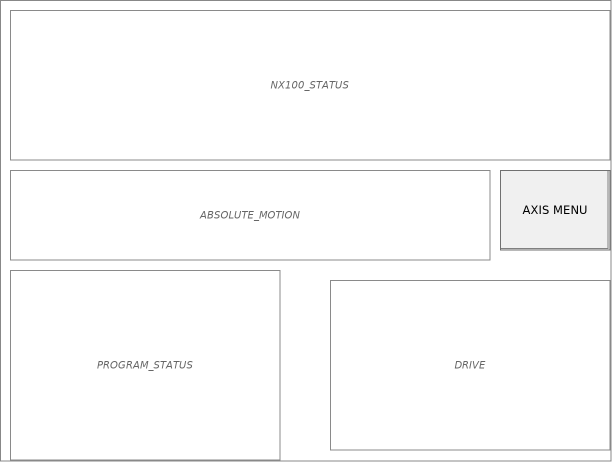
VISUALIZATION TC_VISU  // 612x462
    Frame (10,170 480x90)
        shows ABSOLUTE_MOTION()
    Frame (330,280 280x170)
        shows DRIVE()
    Button (500,170 110x80), "AXIS MENU"
        OnMouseUp: change screen: AXIS
    Frame (10,10 600x150)
        shows NX100_STATUS()
    Frame (10,270 270x190)
        shows PROGRAM_STATUS()
END_VISUALIZATION

(* stored: Version 1.1.0.1, ProductVersion 3.1.4024.16
   Visu TC_VISU: Id {18ea0383-8a6f-45cd-a2c7-3dd0270ce4c8} *)
